(* IEC 61131-3 sources: twincat-st/tests/fixtures/positive, 6 files *)

(* ---- FB_ConditionalCalls.st ---- *)
// X12: a timer, a trigger and a motion block each called only inside a branch.
// CP7: the motion block's Error is never read, nor is the house FB's bError.
// CP12: the valve output is written from the body and from a method.
FUNCTION_BLOCK FB_Device
VAR_INPUT
    bExecute : BOOL;
END_VAR
VAR_OUTPUT
    bDone    : BOOL;
    bError   : BOOL;
END_VAR
bDone := bExecute;
bError := FALSE;
END_FUNCTION_BLOCK

FUNCTION_BLOCK FB_ConditionalCalls
VAR_INPUT
    bStart   : BOOL;
    bSensor  : BOOL;
    fPos     : LREAL;    // mm
END_VAR
VAR_OUTPUT
    bBusy    : BOOL;
END_VAR
VAR
    eStep    : E_Step;
    tonWait  : TON;
    fbEdge   : R_TRIG;
    fbMove   : MC_MoveAbsolute;
    fbDevice : FB_Device;
    axisX    : AXIS_REF;
    qbValve AT %Q* : BOOL;
END_VAR
CASE eStep OF
    E_Step.Idle:
        IF bStart THEN
            eStep := E_Step.Wait;
        END_IF
    E_Step.Wait:
        tonWait(IN := TRUE, PT := T#2S);
        fbEdge(CLK := bSensor);
        IF tonWait.Q OR fbEdge.Q THEN
            eStep := E_Step.Move;
        END_IF
    E_Step.Move:
        fbMove(Axis := axisX, Execute := TRUE, Position := fPos, Velocity := 50.0);
        IF fbMove.Done THEN
            eStep := E_Step.Idle;
        END_IF
    E_Step.Error:
        eStep := E_Step.Idle;
ELSE
    eStep := E_Step.Error;
END_CASE
fbDevice(bExecute := bStart);
qbValve := eStep = E_Step.Move;
bBusy := fbDevice.bDone;
END_FUNCTION_BLOCK

METHOD CloseValve
qbValve := FALSE;
END_METHOD

(* ---- FB_LatchedCompare.st ---- *)
// CP8 skips change detection against a latched copy (fTarget <> fSetpoint), but
// a measured position compared exactly with that same target was never copied
// from it and must still fire. A field test found both shapes side by side.
FUNCTION_BLOCK FB_LatchedCompare
VAR_INPUT
  fSetpoint  : LREAL;  // [mm]
  fActPos    : LREAL;  // [mm] from the axis
  bStart     : BOOL;
END_VAR
VAR_OUTPUT
  bSetpointChanged : BOOL;
  bInPosition      : BOOL;
END_VAR
VAR
  fTarget    : LREAL;  // [mm] setpoint latched at start
END_VAR
IF bStart THEN
  fTarget := fSetpoint;
END_IF
bSetpointChanged := (fTarget <> fSetpoint);
bInPosition := (fActPos = fTarget);
END_FUNCTION_BLOCK

(* ---- FB_LevelExecute.st ---- *)
// X11: both moves are fed from a level. The first is the field test's B2b prompt
// as given; the second is what an agent delivered next to it. Each starts once,
// on its first rising edge, and never again while the expression stays TRUE.
FUNCTION_BLOCK FB_LevelExecute
VAR_INPUT
    bAutoMode : BOOL;
    bAtHome   : BOOL;
    bPicked   : BOOL;
    fPickPos  : LREAL;
    fPlacePos : LREAL;
    fVelo     : LREAL;
END_VAR
VAR
    fbMovePick  : MC_MoveAbsolute;
    fbMovePlace : MC_MoveAbsolute;
    axisX       : AXIS_REF;
END_VAR
fbMovePick(Axis := axisX, Execute := bAutoMode AND bAtHome, Position := fPickPos, Velocity := fVelo);
fbMovePlace.Execute := bAutoMode AND bPicked AND NOT fbMovePick.Busy;
fbMovePlace(Axis := axisX, Position := fPlacePos, Velocity := fVelo);
END_FUNCTION_BLOCK

(* ---- FB_NestedGuardTimer.st ---- *)
// X12: neither guard leaves the timer alone. 'OR NOT bIn' nested under 'bEnable
// AND (...)' is never entered with bEnable FALSE, so fbTimer is never reset; and a
// reference check joined with a run flag is a state branch, not a reference guard.
FUNCTION_BLOCK FB_NestedGuardTimer
VAR_INPUT
    bEnable     : BOOL;
    bUseTimeout : BOOL;
    bIn         : BOOL;
    tTimeout    : TIME;
END_VAR
VAR_IN_OUT
    refCfg : ST_TimerCfg;
END_VAR
VAR_OUTPUT
    bTimedOut : BOOL;
    bInfo     : BOOL;
END_VAR
VAR
    fbTimer : TON;
    fbCheck : TON;
    rCfg    : REFERENCE TO ST_TimerCfg;
END_VAR
rCfg REF= refCfg;
IF bEnable AND (bUseTimeout OR NOT bIn) THEN
    fbTimer(IN := bIn, PT := tTimeout);
END_IF
IF __ISVALIDREF(rCfg) AND bEnable THEN
    fbCheck(IN := bIn, PT := rCfg.tInfo);
END_IF
bTimedOut := fbTimer.Q;
bInfo := fbCheck.Q;
END_FUNCTION_BLOCK

(* ---- FB_PragmaDecl.st ---- *)
// A declaration behind a pragma line is a declaration. The parser used to drop
// each one, so no rule saw it. nHidden is never used (CP24, reported on its own
// line, not the pragma's); nStep is marked TcRetain and steps its CASE (X13).
FUNCTION_BLOCK FB_PragmaDecl
VAR_INPUT
    bStart : BOOL;
END_VAR
VAR_OUTPUT
    bError : BOOL;
END_VAR
VAR
    {attribute 'hide'}
    nHidden : INT;
    {attribute 'TcRetain'}
    nStep : INT;
END_VAR
CASE nStep OF
    0:  IF bStart THEN nStep := 10; END_IF
    10: IF NOT bStart THEN nStep := 0; END_IF
    99: bError := TRUE;
        IF NOT bStart THEN bError := FALSE; nStep := 0; END_IF
ELSE
    nStep := 99;
END_CASE
END_FUNCTION_BLOCK

(* ---- FB_RemanentStep.st ---- *)
// X13: a state machine's step declared remanent, in both forms Haiku wrote in the
// homed-survives-restart eval: a VAR RETAIN block, and the qualifier after the type.
// X14: that second form, which is not where IEC 61131-3 puts the qualifier.
FUNCTION_BLOCK FB_RemanentStep
VAR_INPUT
    bStart  : BOOL;
    bAtHome : BOOL;
END_VAR
VAR_OUTPUT
    bHomed : BOOL;
    bError : BOOL;
END_VAR
VAR RETAIN
    nStep : INT;
END_VAR
VAR
    nPhase : INT PERSISTENT;
END_VAR
CASE nStep OF
    0:  IF bStart THEN nStep := 10; END_IF
    10: IF bAtHome THEN bHomed := TRUE; nStep := 20; END_IF
    20: IF NOT bStart THEN bHomed := FALSE; nStep := 0; END_IF
    99: bError := TRUE;
        IF NOT bStart THEN bError := FALSE; nStep := 0; END_IF
ELSE
    nStep := 99;
END_CASE
CASE nPhase OF
    0: IF bHomed THEN nPhase := 1; END_IF
    1: IF NOT bHomed THEN nPhase := 0; END_IF
ELSE
    nPhase := 0;
END_CASE
END_FUNCTION_BLOCK
